Staubli VAL3: setLabelValue.pgx

public program setLabelValue(num x_nType)
  local num l_nSize
  local num l_i
  local string l_slabel
  local num l_nSize1
begin

  call getSize(l_nSize,l_nSize1)
  //
  switch x_nType
    case 0
      for l_i = 0 to l_nSize-1
        sLabel[l_i]=toString("",l_i+16*nPageIndex)+".dIn["+toString("",l_i+16*nPageIndex)+"]"
        sComment[l_i]=io:dInItem[l_i+16*nPageIndex].sComment
      endFor
    break
    case 1
      for l_i = 0 to l_nSize-1
        sLabel[l_i]=toString("",l_i+16*nPageIndex)+".dOut["+toString("",l_i+16*nPageIndex)+"]"
        sComment[l_i]=io:dOutItem[l_i+16*nPageIndex].sComment
      endFor
    break
    case 2
      for l_i = 0 to l_nSize1-1
        sLabel[l_i]=toString("",l_i+16*nPageIndex)+".aIn["+toString("",l_i+16*nPageIndex)+"]"
        sComment[l_i]=io:aInItem[l_i+16*nPageIndex].sComment
      endFor
    break
    case 3
      for l_i = 0 to l_nSize1-1
        sLabel[l_i]=toString("",l_i+16*nPageIndex)+".aOut["+toString("",l_i+16*nPageIndex)+"]"
        sComment[l_i]=io:aOutItem[l_i+16*nPageIndex].sComment
      endFor

    break
  endSwitch

end
